{attribute 'linkalways'}
{attribute 'no_explicit_call' := 'Use the methods of this class'}
{attribute 'enable_dynamic_creation'}
FUNCTION_BLOCK WheelOdometry IMPLEMENTS I_PoseSource
VAR
	drive : I_DifferentialDrive;
	kinematics : DiffDriveKinematics;
	_pose : Pose2D;
	lastLeftInM : LREAL;
	lastRightInM : LREAL;
END_VAR

METHOD Connect
VAR_INPUT
	differentialDrive : I_DifferentialDrive;
END_VAR
drive := differentialDrive;
END_METHOD

METHOD Execute
VAR
	leftInM : LREAL;
	rightInM : LREAL;
	motion : BodyMotion;
	midHeadingInRad : LREAL;
END_VAR
leftInM := drive.LeftWheelPositionInM;
rightInM := drive.RightWheelPositionInM;

motion := kinematics.ToBodyMotion(leftDeltaInM := leftInM - lastLeftInM, rightDeltaInM := rightInM - lastRightInM);
lastLeftInM := leftInM;
lastRightInM := rightInM;

midHeadingInRad := _pose.thetaInRad + motion.headingChangeInRad / 2.0;
_pose.x := _pose.x + motion.distanceInM * COS(midHeadingInRad);
_pose.y := _pose.y + motion.distanceInM * SIN(midHeadingInRad);
_pose.thetaInRad := _pose.thetaInRad + motion.headingChangeInRad;

IF _pose.thetaInRad > PI THEN
	_pose.thetaInRad := _pose.thetaInRad - 2.0 * PI;
ELSIF _pose.thetaInRad <= -PI THEN
	_pose.thetaInRad := _pose.thetaInRad + 2.0 * PI;
END_IF
END_METHOD

PROPERTY Pose : Pose2D
GET
Pose := _pose;
END_GET
END_PROPERTY

METHOD Reset
VAR_INPUT
	pose : Pose2D;
END_VAR
_pose := pose;

lastLeftInM := drive.LeftWheelPositionInM;
lastRightInM := drive.RightWheelPositionInM;
END_METHOD

END_FUNCTION_BLOCK

(* stored: Version 1.1.0.1
   POU WheelOdometry: Id {0383d384-f1af-5157-a3ab-6329c1f8f315}, SpecialFunc None
   Method Connect: Id {9586be9c-1b18-592a-ac72-9a0cd025658c}
   Method Execute: Id {2ece7e54-0fcd-5291-83ae-9ff6c29c3813}
   Property Pose: Id {7cb73c2f-8b0e-5f16-82ed-16a14c60a740}
   Get Get: Id {0a0650ae-20a5-5470-a202-fff7e5873f72}
   Method Reset: Id {eac72228-2ae7-507b-bd27-7b6833793730} *)
